(* Logix 5000 project; controller R400_500_XLS vendor 1 type 14 code 216 rev 31.11; software revision 31.01; part 6 of 32 *)
(* tags used below, declared in another part *)
   Abort1 : DINT;   // Not Used
   Alarm : SINT;   // Wait 3 seconds
   AlarmAcked : BOOL;   // Alarm has been acked
   Ashutdown : SINT;   // Not Used
   bAlrm : BOOL[64];
   CycleSequence : UDT_CYCLE_SEQUENCE;
   Drain_RcvryTnk_with_Sump : DINT;   // 0 = Close Recovery Tank Drain Valve 1 = Open Recovery Tank Drain Valve
   DrnSmp : DINT;
   DRYING : DINT;   // Drying id number
   M : DINT[5];   // Memory Bits
   OneShot : DINT[1];
   ONS_FC25 : DINT;
   PrimeChemPmp : SINT;   // Prime chemical pumps activation bits
   Rcvry_Tnk_Tmp : REAL;   // Water Temperature of the Heat Recovery Tank
   Service : DINT[2];   // Unused Service Mode Memory Bit
   Shutdown : SINT;   // Shutdown sequence steps
   Shutdown_Tran : SINT;   // Shutdown sequence transitions
   Tmr : TIMER[107];
   AlarmMsg : STRING;   // Message of the alarm from the HMI Do not delete this tag
   AlarmTrigger : INT;   // Triggers the alarm screen if different of 0
   bAcceptRejectRecorded : BOOL;   // Cycle Accept/Reject Recorded By User
   Cfg_10_Modules : BOOL;   // Chassis is configured 10 slots
   Cfg_11_Modules : BOOL;
   Current_Screen : DINT;
   CycleUsage : UDT_CYCLE_USAGE[50];
   EmailSMSInt : INT[8];   // Email & SMS Notification Integer
   I_Ld_Dr_Cls_Sw : BOOL;   // Load door close
   I_Pw_Tnk_Lvl_Sw : BOOL;   // Pure water tank level switch
   I_Unld_Dr_Cls_Sw : BOOL;   // Unload door close
   MaintainCloseLd : BOOL;
   MaintainCloseUnld : BOOL;
   MaintainOpenLd : BOOL;
   MaintainOpenUnld : BOOL;
   msg : BOOL[512];
   Msg_Shutdown : SINT;
   Q_Chm_1 : BOOL;   // Chemical pump #1
   Q_Chm_2 : BOOL;   // Chemical pump #2
   Q_Chm_3 : BOOL;   // Chemical pump #3
   Q_Chm_4 : BOOL;   // Chemical pump #4
   Q_Ht_Rcvry_Tnk_Drn_Vlve : BOOL;   // Heat recovery tank drian valve
   Screen_Ctrl : DINT;   // PLC Screen Request
   Tpb : DINT[11];
   TpbImage : DINT[11];
   Unit : Hrdwre;   // Unit Configuration
(* MainProgram, continued *)

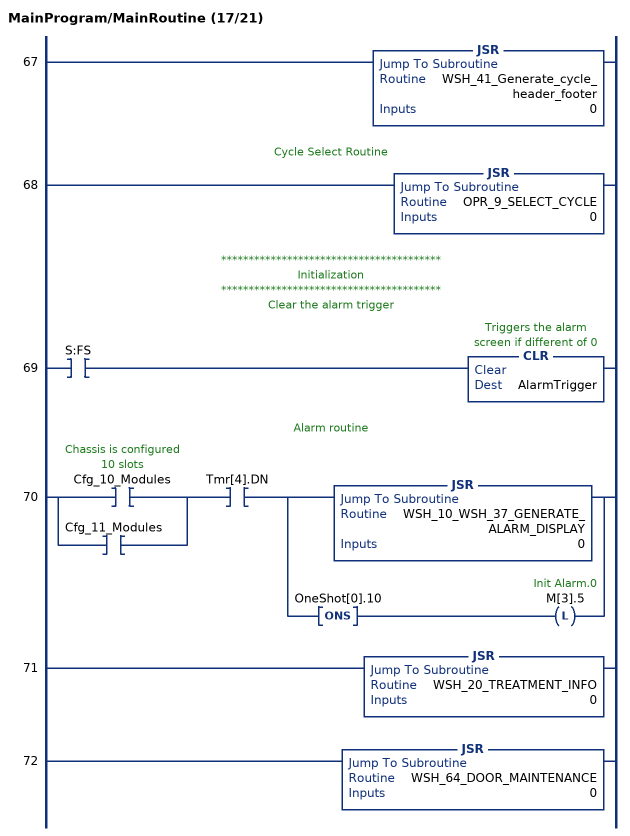
   [picture p68: MainProgram/MainRoutine rungs 67-72]
   67: JSR(WSH_41_Generate_cycle_header_footer,0);
   // Cycle Select Routine
   68: JSR(OPR_9_SELECT_CYCLE,0);
   // ****************************************
   // Initialization
   // ****************************************
   // Clear the alarm trigger
   69: XIC(S:FS)CLR(AlarmTrigger);
   // Alarm routine
   70: [XIC(Cfg_10_Modules) ,XIC(Cfg_11_Modules) ]XIC(Tmr[4].DN)[JSR(WSH_10_WSH_37_GENERATE_ALARM_DISPLAY,0) ,ONS(OneShot[0].10) OTL(M[3].5) ];
   71: JSR(WSH_20_TREATMENT_INFO,0);
   72: JSR(WSH_64_DOOR_MAINTENANCE,0);
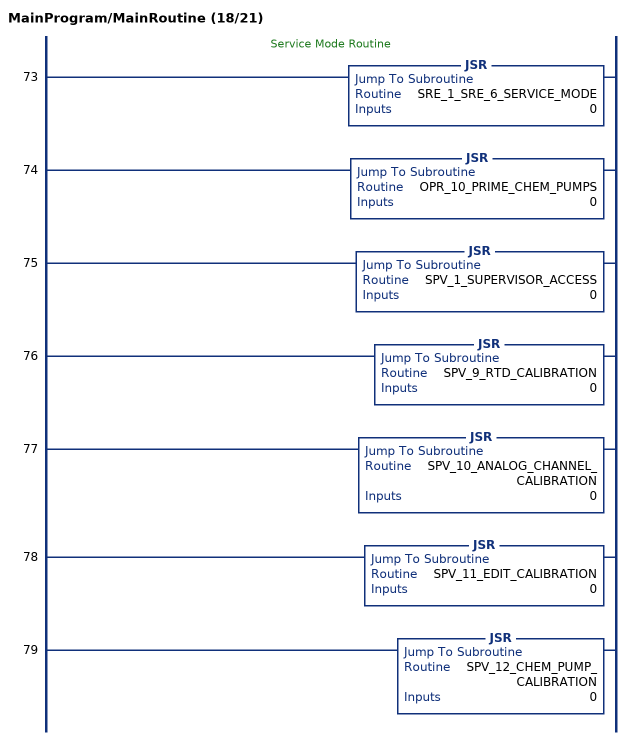
   // Service Mode Routine
   73: JSR(SRE_1_SRE_6_SERVICE_MODE,0);
   74: JSR(OPR_10_PRIME_CHEM_PUMPS,0);
   75: JSR(SPV_1_SUPERVISOR_ACCESS,0);
   76: JSR(SPV_9_RTD_CALIBRATION,0);
   77: JSR(SPV_10_ANALOG_CHANNEL_CALIBRATION,0);
   78: JSR(SPV_11_EDIT_CALIBRATION,0);
   79: JSR(SPV_12_CHEM_PUMP_CALIBRATION,0);
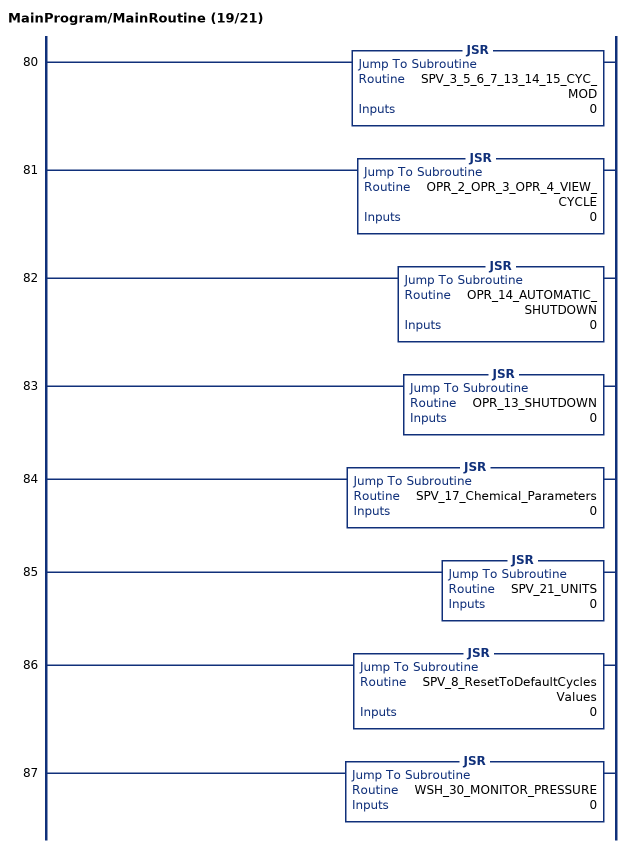
   80: JSR(SPV_3_5_6_7_13_14_15_CYC_MOD,0);
   81: JSR(OPR_2_OPR_3_OPR_4_VIEW_CYCLE,0);
   82: JSR(OPR_14_AUTOMATIC_SHUTDOWN,0);
   83: JSR(OPR_13_SHUTDOWN,0);
   84: JSR(SPV_17_Chemical_Parameters,0);
   85: JSR(SPV_21_UNITS,0);
   86: JSR(SPV_8_ResetToDefaultCyclesValues,0);
   87: JSR(WSH_30_MONITOR_PRESSURE,0);
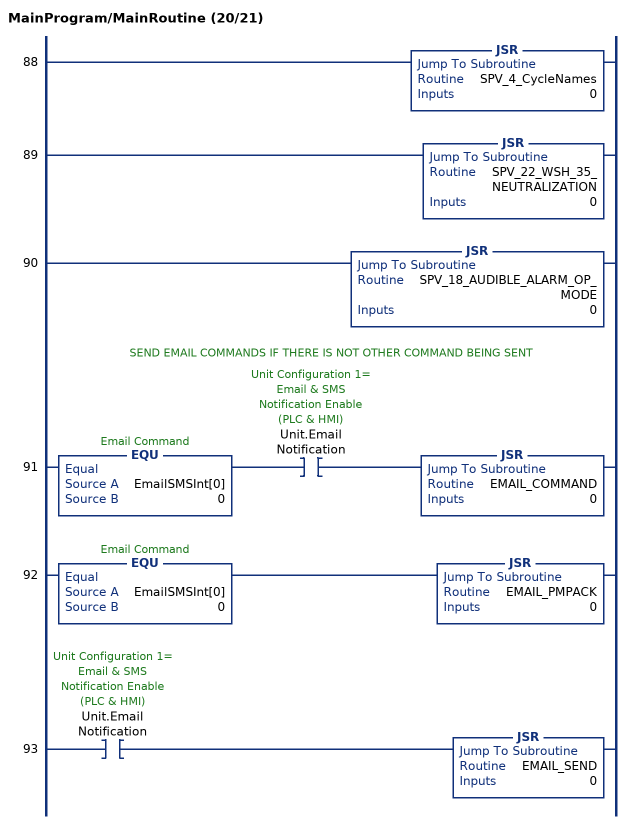
   88: JSR(SPV_4_CycleNames,0);
   89: JSR(SPV_22_WSH_35_NEUTRALIZATION,0);
   90: JSR(SPV_18_AUDIBLE_ALARM_OP_MODE,0);
   // SEND EMAIL COMMANDS IF THERE IS NOT OTHER COMMAND BEING SENT
   91: EQU(EmailSMSInt[0],0)XIC(Unit.EmailNotification)JSR(EMAIL_COMMAND,0);
   92: EQU(EmailSMSInt[0],0)JSR(EMAIL_PMPACK,0);
   93: XIC(Unit.EmailNotification)JSR(EMAIL_SEND,0);
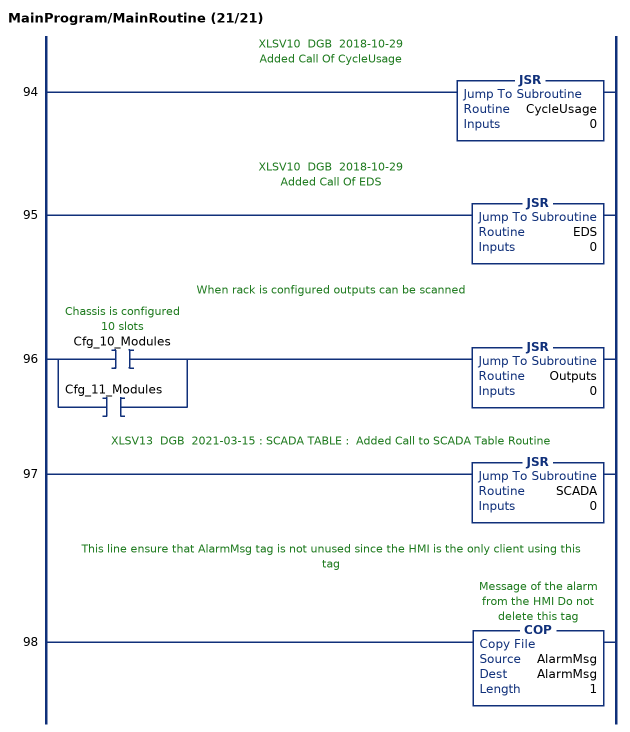
   // XLSV10  DGB  2018-10-29
   // Added Call Of CycleUsage
   94: JSR(CycleUsage,0);
   // XLSV10  DGB  2018-10-29
   // Added Call Of EDS
   95: JSR(EDS,0);
   // When rack is configured outputs can be scanned
   96: [XIC(Cfg_10_Modules) ,XIC(Cfg_11_Modules) ]JSR(Outputs,0);
   // XLSV13  DGB  2021-03-15 : SCADA TABLE :  Added Call to SCADA Table Routine
   97: JSR(SCADA,0);
   // This line ensure that AlarmMsg tag is not unused since the HMI is the only client using this  tag
   98: COP(AlarmMsg,AlarmMsg,1);
END_ROUTINE

ROUTINE OPR_10_PRIME_CHEM_PUMPS   (* ladder *)
// Prime chemical pumps routine
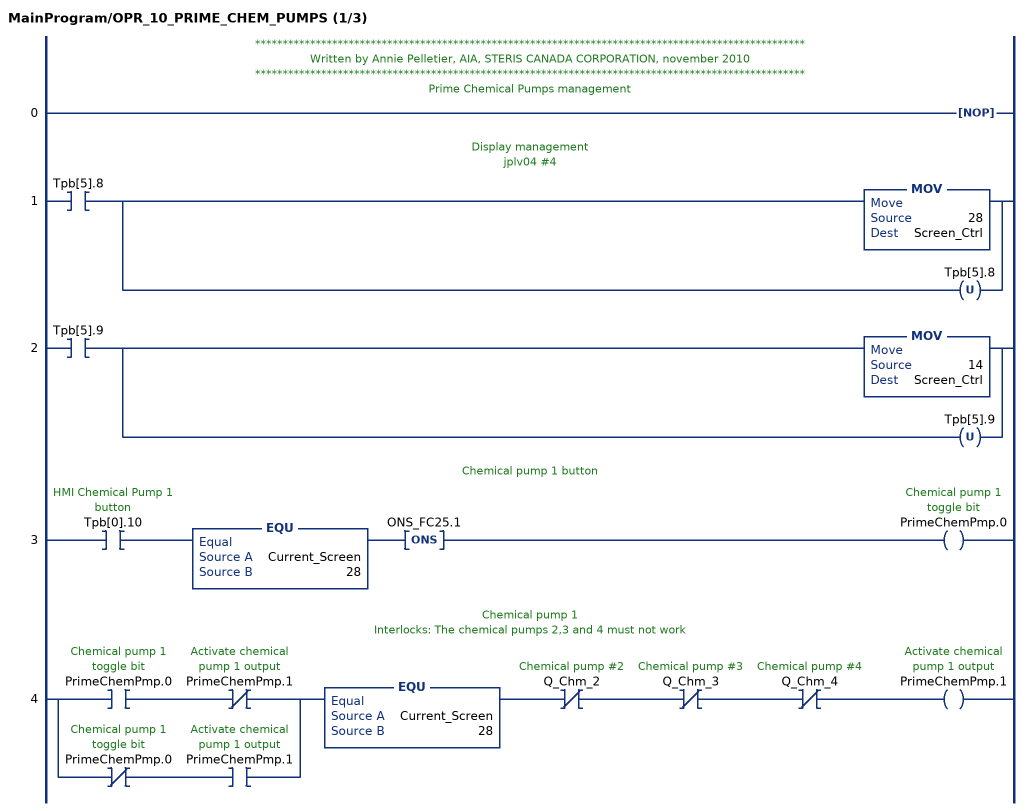
   // ****************************************************************************************************
   // Written by Annie Pelletier, AIA, STERIS CANADA CORPORATION, november 2010
   // ****************************************************************************************************
   // Prime Chemical Pumps management
   0: NOP();
   // Display management
   // jplv04 #4
   1: XIC(Tpb[5].8)[MOV(28,Screen_Ctrl) ,OTU(Tpb[5].8) ];
   2: XIC(Tpb[5].9)[MOV(14,Screen_Ctrl) ,OTU(Tpb[5].9) ];
   // Chemical pump 1 button
   3: XIC(Tpb[0].10)EQU(Current_Screen,28)ONS(ONS_FC25.1)OTE(PrimeChemPmp.0);
   // Chemical pump 1
   // Interlocks: The chemical pumps 2,3 and 4 must not work
   4: [XIC(PrimeChemPmp.0) XIO(PrimeChemPmp.1) ,XIO(PrimeChemPmp.0) XIC(PrimeChemPmp.1) ]EQU(Current_Screen,28)XIO(Q_Chm_2)XIO(Q_Chm_3)XIO(Q_Chm_4)OTE(PrimeChemPmp.1);
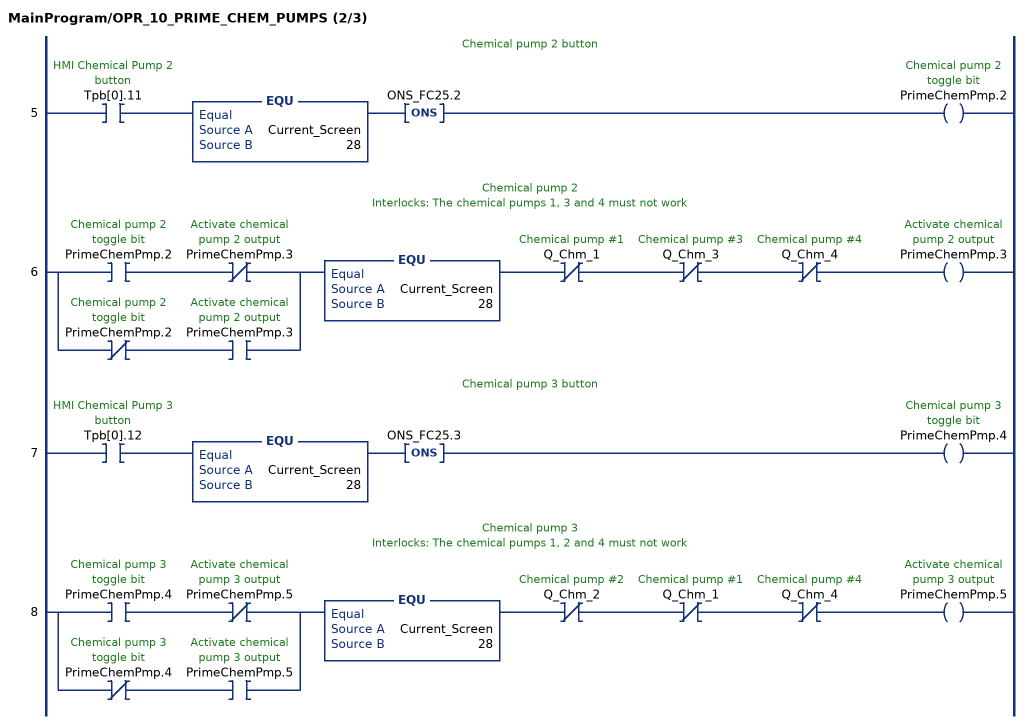
   // Chemical pump 2 button
   5: XIC(Tpb[0].11)EQU(Current_Screen,28)ONS(ONS_FC25.2)OTE(PrimeChemPmp.2);
   // Chemical pump 2
   // Interlocks: The chemical pumps 1, 3 and 4 must not work
   6: [XIC(PrimeChemPmp.2) XIO(PrimeChemPmp.3) ,XIO(PrimeChemPmp.2) XIC(PrimeChemPmp.3) ]EQU(Current_Screen,28)XIO(Q_Chm_1)XIO(Q_Chm_3)XIO(Q_Chm_4)OTE(PrimeChemPmp.3);
   // Chemical pump 3 button
   7: XIC(Tpb[0].12)EQU(Current_Screen,28)ONS(ONS_FC25.3)OTE(PrimeChemPmp.4);
   // Chemical pump 3
   // Interlocks: The chemical pumps 1, 2 and 4 must not work
   8: [XIC(PrimeChemPmp.4) XIO(PrimeChemPmp.5) ,XIO(PrimeChemPmp.4) XIC(PrimeChemPmp.5) ]EQU(Current_Screen,28)XIO(Q_Chm_2)XIO(Q_Chm_1)XIO(Q_Chm_4)OTE(PrimeChemPmp.5);
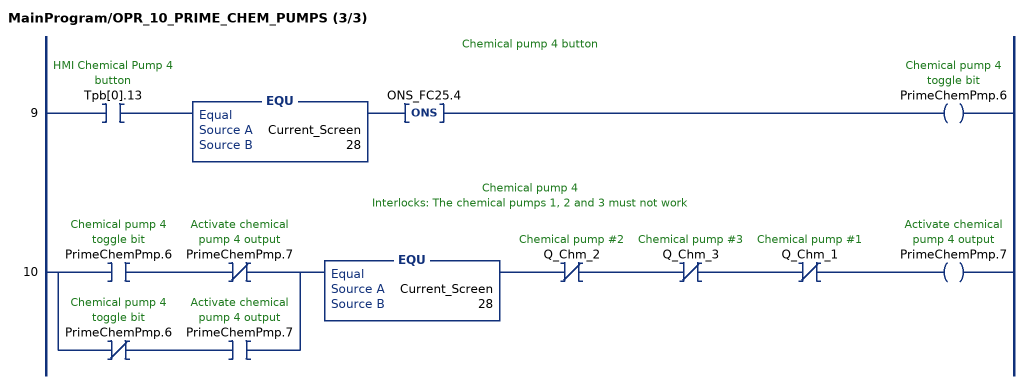
   // Chemical pump 4 button
   9: XIC(Tpb[0].13)EQU(Current_Screen,28)ONS(ONS_FC25.4)OTE(PrimeChemPmp.6);
   // Chemical pump 4
   // Interlocks: The chemical pumps 1, 2 and 3 must not work
   10: [XIC(PrimeChemPmp.6) XIO(PrimeChemPmp.7) ,XIO(PrimeChemPmp.6) XIC(PrimeChemPmp.7) ]EQU(Current_Screen,28)XIO(Q_Chm_2)XIO(Q_Chm_3)XIO(Q_Chm_1)OTE(PrimeChemPmp.7);
END_ROUTINE

ROUTINE OPR_13_SHUTDOWN   (* ladder *)
// This routine manage the washer's shutdown
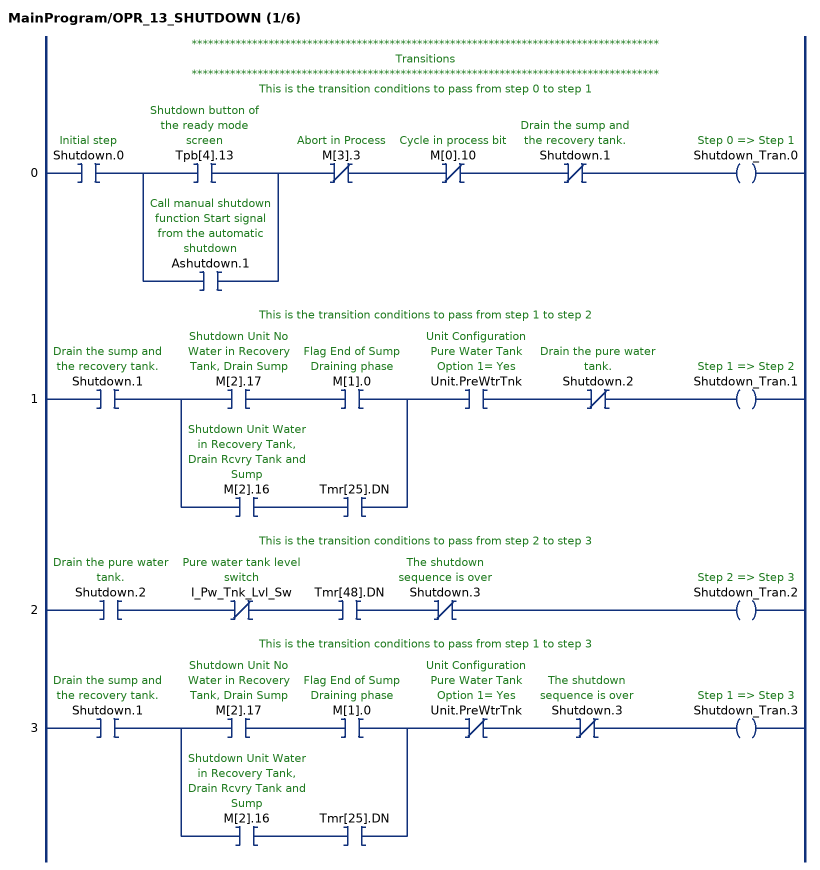
   // *************************************************************************************
   // Transitions
   // *************************************************************************************
   // This is the transition conditions to pass from step 0 to step 1
   0: XIC(Shutdown.0)[XIC(Tpb[4].13) ,XIC(Ashutdown.1) ]XIO(M[3].3)XIO(M[0].10)XIO(Shutdown.1)OTE(Shutdown_Tran.0);
   // This is the transition conditions to pass from step 1 to step 2
   1: XIC(Shutdown.1)[XIC(M[2].17) XIC(M[1].0) ,XIC(M[2].16) XIC(Tmr[25].DN) ]XIC(Unit.PreWtrTnk)XIO(Shutdown.2)OTE(Shutdown_Tran.1);
   // This is the transition conditions to pass from step 2 to step 3
   2: XIC(Shutdown.2)XIO(I_Pw_Tnk_Lvl_Sw)XIC(Tmr[48].DN)XIO(Shutdown.3)OTE(Shutdown_Tran.2);
   // This is the transition conditions to pass from step 1 to step 3
   3: XIC(Shutdown.1)[XIC(M[2].17) XIC(M[1].0) ,XIC(M[2].16) XIC(Tmr[25].DN) ]XIO(Unit.PreWtrTnk)XIO(Shutdown.3)OTE(Shutdown_Tran.3);
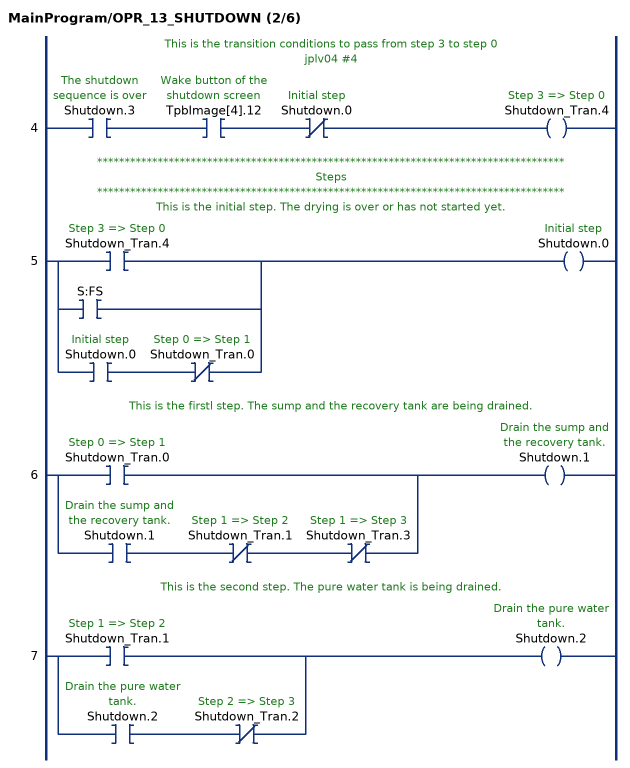
   // This is the transition conditions to pass from step 3 to step 0
   // jplv04 #4
   4: XIC(Shutdown.3)XIC(TpbImage[4].12)XIO(Shutdown.0)OTE(Shutdown_Tran.4);
   // *************************************************************************************
   // Steps
   // *************************************************************************************
   // This is the initial step. The drying is over or has not started yet.
   5: [XIC(Shutdown_Tran.4) ,XIC(S:FS) ,XIC(Shutdown.0) XIO(Shutdown_Tran.0) ]OTE(Shutdown.0);
   // This is the firstl step. The sump and the recovery tank are being drained.
   6: [XIC(Shutdown_Tran.0) ,XIC(Shutdown.1) XIO(Shutdown_Tran.1) XIO(Shutdown_Tran.3) ]OTE(Shutdown.1);
   // This is the second step. The pure water tank is being drained.
   7: [XIC(Shutdown_Tran.1) ,XIC(Shutdown.2) XIO(Shutdown_Tran.2) ]OTE(Shutdown.2);
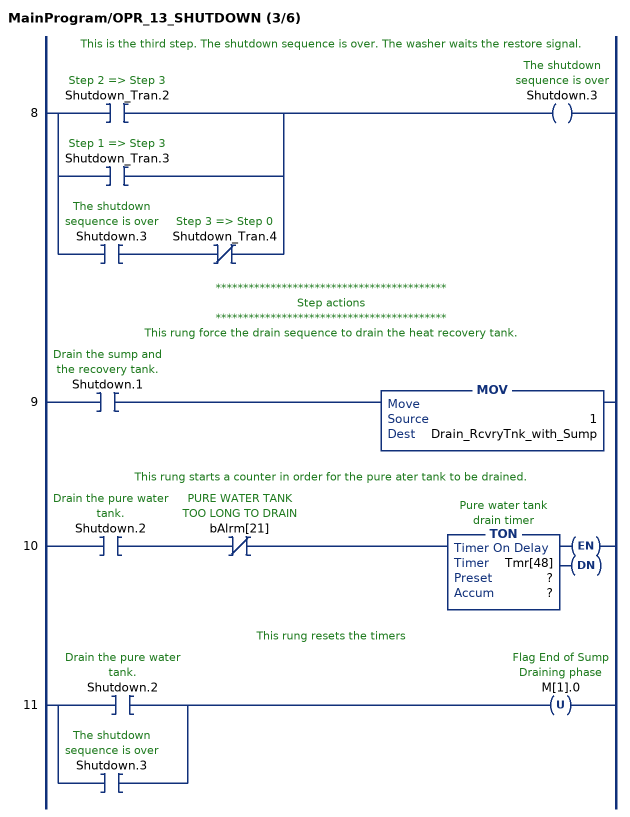
   // This is the third step. The shutdown sequence is over. The washer waits the restore signal.
   8: [XIC(Shutdown_Tran.2) ,XIC(Shutdown_Tran.3) ,XIC(Shutdown.3) XIO(Shutdown_Tran.4) ]OTE(Shutdown.3);
   // ******************************************
   // Step actions
   // ******************************************
   // This rung force the drain sequence to drain the heat recovery tank.
   9: XIC(Shutdown.1)MOV(1,Drain_RcvryTnk_with_Sump);
   // This rung starts a counter in order for the pure ater tank to be drained.
   10: XIC(Shutdown.2)XIO(bAlrm[21])TON(Tmr[48],?,?);
   // This rung resets the timers
   11: [XIC(Shutdown.2) ,XIC(Shutdown.3) ]OTU(M[1].0);
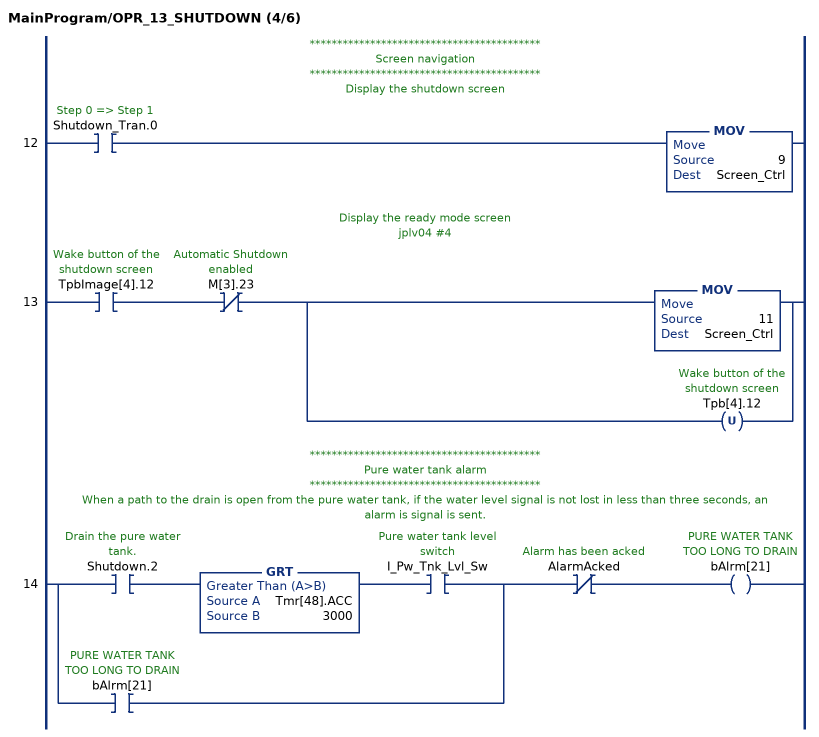
   // ******************************************
   // Screen navigation
   // ******************************************
   // Display the shutdown screen
   12: XIC(Shutdown_Tran.0)MOV(9,Screen_Ctrl);
   // Display the ready mode screen
   // jplv04 #4
   13: XIC(TpbImage[4].12)XIO(M[3].23)[MOV(11,Screen_Ctrl) ,OTU(Tpb[4].12) ];
   // ******************************************
   // Pure water tank alarm
   // ******************************************
   // When a path to the drain is open from the pure water tank, if the water level signal is not lost in less than three seconds, an alarm is signal is sent.
   14: [XIC(Shutdown.2) GRT(Tmr[48].ACC,3000) XIC(I_Pw_Tnk_Lvl_Sw) ,XIC(bAlrm[21]) ]XIO(AlarmAcked)OTE(bAlrm[21]);
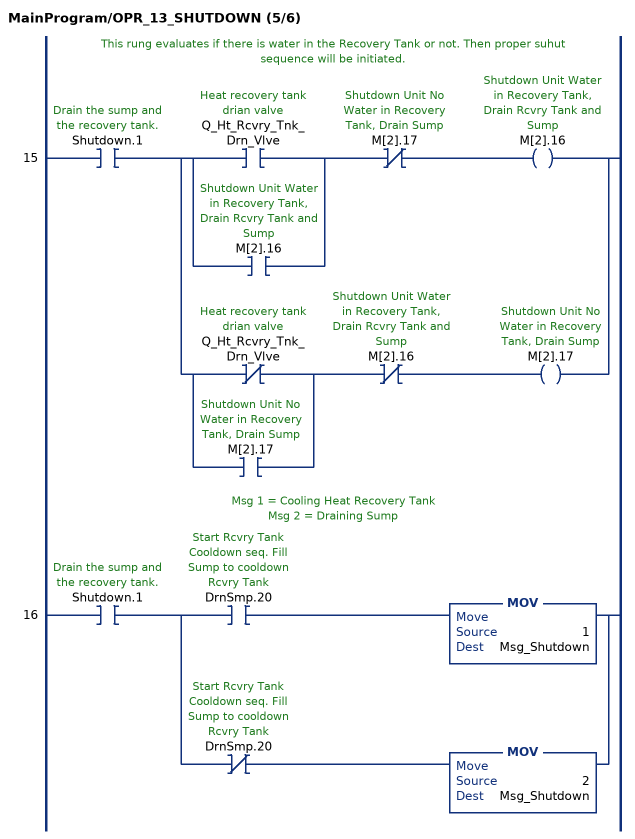
   // This rung evaluates if there is water in the Recovery Tank or not. Then proper suhut sequence will be initiated.
   15: XIC(Shutdown.1)[[XIC(Q_Ht_Rcvry_Tnk_Drn_Vlve) ,XIC(M[2].16) ] XIO(M[2].17) OTE(M[2].16) ,[XIO(Q_Ht_Rcvry_Tnk_Drn_Vlve) ,XIC(M[2].17) ] XIO(M[2].16) OTE(M[2].17) ];
   // Msg 1 = Cooling Heat Recovery Tank
   // Msg 2 = Draining Sump
   16: XIC(Shutdown.1)[XIC(DrnSmp.20) MOV(1,Msg_Shutdown) ,XIO(DrnSmp.20) MOV(2,Msg_Shutdown) ];
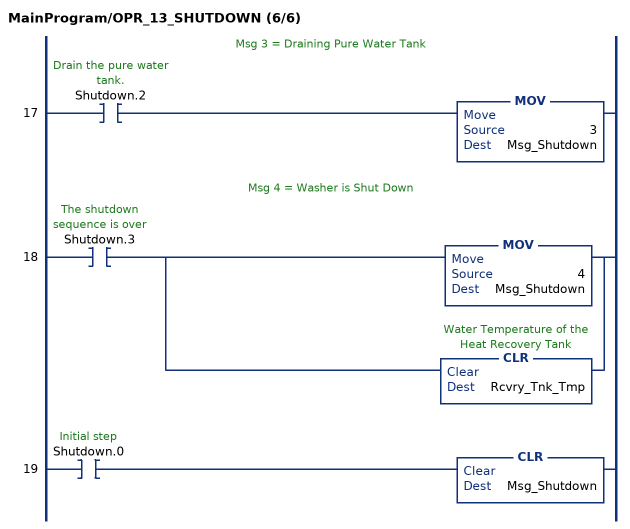
   // Msg 3 = Draining Pure Water Tank
   17: XIC(Shutdown.2)MOV(3,Msg_Shutdown);
   // Msg 4 = Washer is Shut Down
   18: XIC(Shutdown.3)[MOV(4,Msg_Shutdown) ,CLR(Rcvry_Tnk_Tmp) ];
   19: XIC(Shutdown.0)CLR(Msg_Shutdown);
END_ROUTINE

ROUTINE OPR_14_AUTOMATIC_SHUTDOWN   (* ladder *)
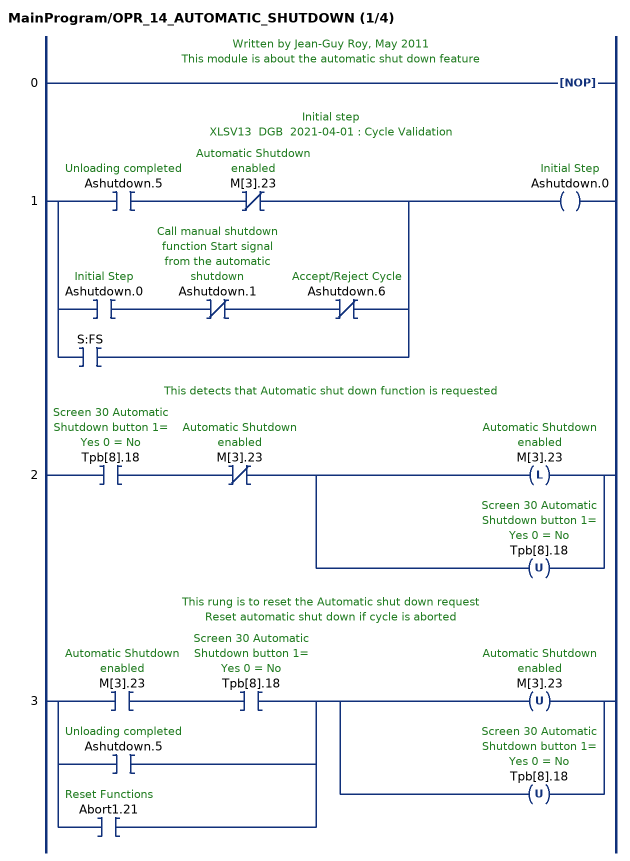
   // Written by Jean-Guy Roy, May 2011
   // This module is about the automatic shut down feature
   0: NOP();
   // Initial step
   // XLSV13  DGB  2021-04-01 : Cycle Validation
   1: [XIC(Ashutdown.5) XIO(M[3].23) ,XIC(Ashutdown.0) XIO(Ashutdown.1) XIO(Ashutdown.6) ,XIC(S:FS) ]OTE(Ashutdown.0);
   // This detects that Automatic shut down function is requested
   2: XIC(Tpb[8].18)XIO(M[3].23)[OTL(M[3].23) ,OTU(Tpb[8].18) ];
   // This rung is to reset the Automatic shut down request
   // Reset automatic shut down if cycle is aborted
   3: [XIC(M[3].23) XIC(Tpb[8].18) ,XIC(Ashutdown.5) ,XIC(Abort1.21) ][OTU(M[3].23) ,OTU(Tpb[8].18) ];
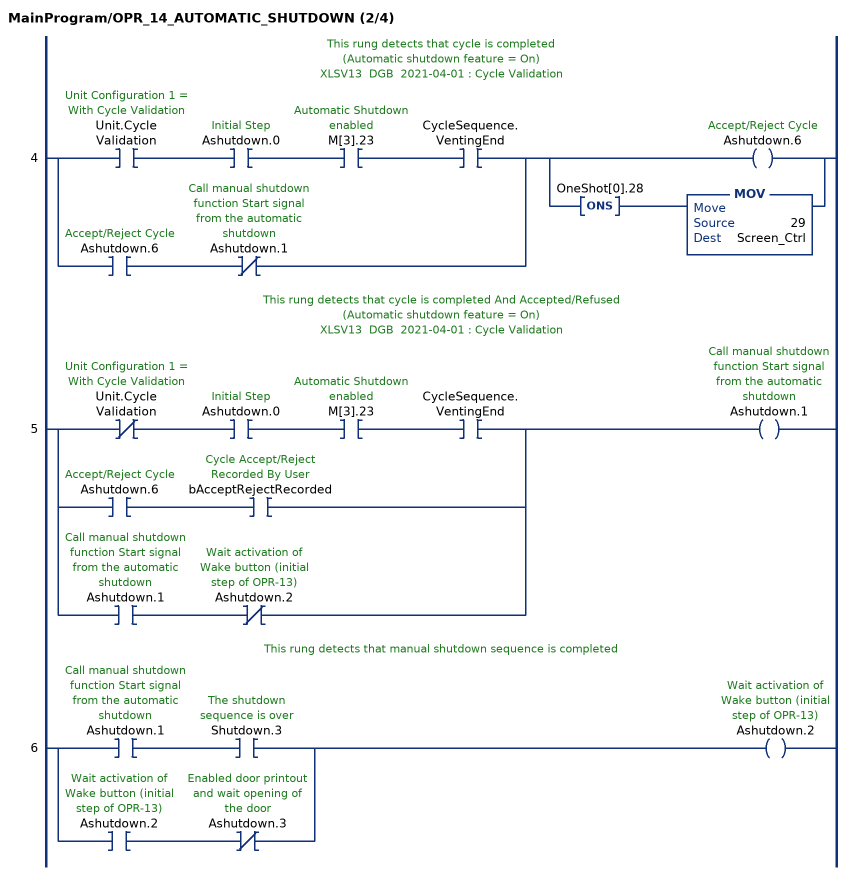
   // This rung detects that cycle is completed
   // (Automatic shutdown feature = On)
   // XLSV13  DGB  2021-04-01 : Cycle Validation
   4: [XIC(Unit.CycleValidation) XIC(Ashutdown.0) XIC(M[3].23) XIC(CycleSequence.VentingEnd) ,XIC(Ashutdown.6) XIO(Ashutdown.1) ][OTE(Ashutdown.6) ,ONS(OneShot[0].28) MOV(29,Screen_Ctrl) ];
   // This rung detects that cycle is completed And Accepted/Refused
   // (Automatic shutdown feature = On)
   // XLSV13  DGB  2021-04-01 : Cycle Validation
   5: [XIO(Unit.CycleValidation) XIC(Ashutdown.0) XIC(M[3].23) XIC(CycleSequence.VentingEnd) ,XIC(Ashutdown.6) XIC(bAcceptRejectRecorded) ,XIC(Ashutdown.1) XIO(Ashutdown.2) ]OTE(Ashutdown.1);
   // This rung detects that manual shutdown sequence is completed
   6: [XIC(Ashutdown.1) XIC(Shutdown.3) ,XIC(Ashutdown.2) XIO(Ashutdown.3) ]OTE(Ashutdown.2);
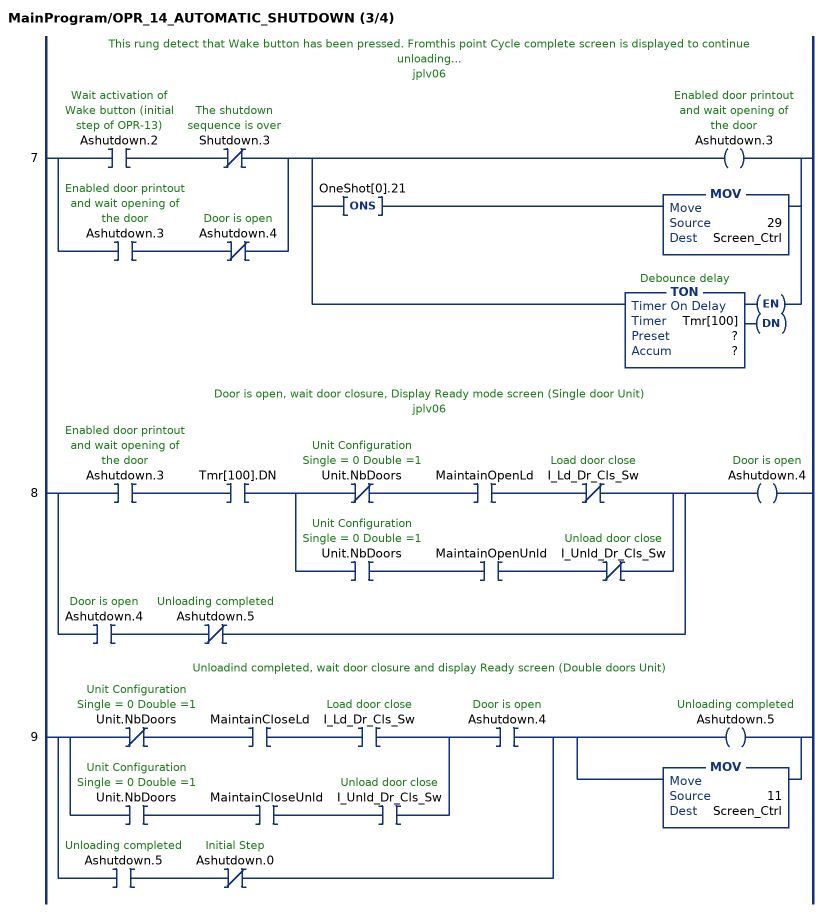
   // This rung detect that Wake button has been pressed. Fromthis point Cycle complete screen is displayed to continue unloading...
   // jplv06
   7: [XIC(Ashutdown.2) XIO(Shutdown.3) ,XIC(Ashutdown.3) XIO(Ashutdown.4) ][OTE(Ashutdown.3) ,ONS(OneShot[0].21) MOV(29,Screen_Ctrl) ,TON(Tmr[100],?,?) ];
   // Door is open, wait door closure, Display Ready mode screen (Single door Unit)
   // jplv06
   8: [XIC(Ashutdown.3) XIC(Tmr[100].DN) [XIO(Unit.NbDoors) XIC(MaintainOpenLd) XIO(I_Ld_Dr_Cls_Sw) ,XIC(Unit.NbDoors) XIC(MaintainOpenUnld) XIO(I_Unld_Dr_Cls_Sw) ] ,XIC(Ashutdown.4) XIO(Ashutdown.5) ]OTE(Ashutdown.4);
   // Unloadind completed, wait door closure and display Ready screen (Double doors Unit)
   9: [[XIO(Unit.NbDoors) XIC(MaintainCloseLd) XIC(I_Ld_Dr_Cls_Sw) ,XIC(Unit.NbDoors) XIC(MaintainCloseUnld) XIC(I_Unld_Dr_Cls_Sw) ] XIC(Ashutdown.4) ,XIC(Ashutdown.5) XIO(Ashutdown.0) ][OTE(Ashutdown.5) ,MOV(11,Screen_Ctrl) ];
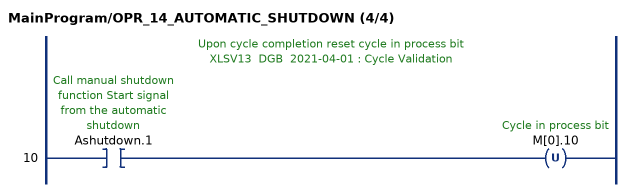
   // Upon cycle completion reset cycle in process bit
   // XLSV13  DGB  2021-04-01 : Cycle Validation
   10: XIC(Ashutdown.1)OTU(M[0].10);
END_ROUTINE
